RoboDK station: T1-instructions.rdk

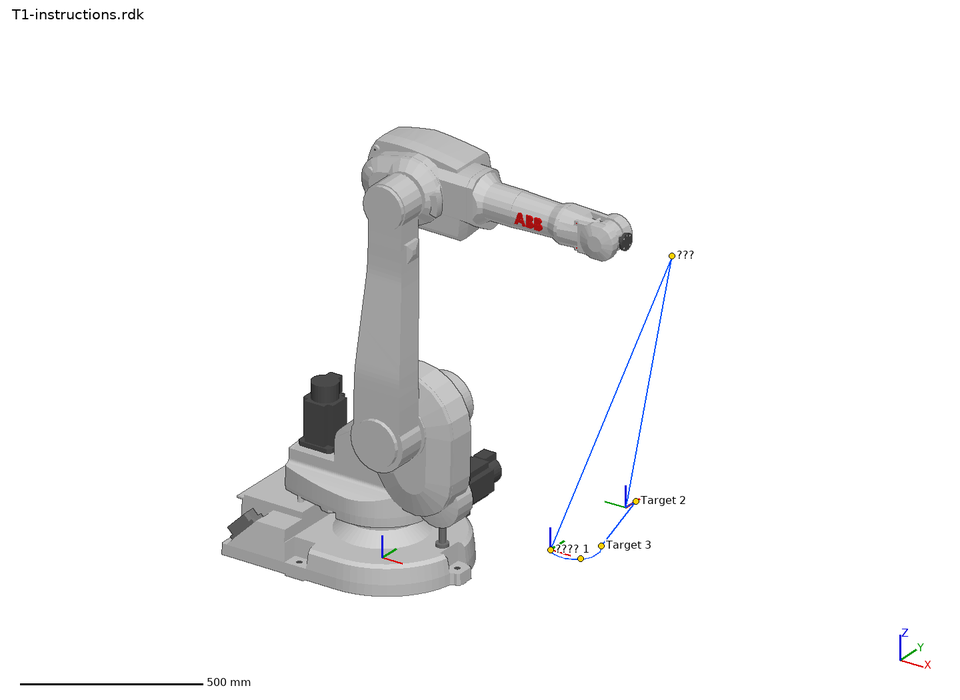
[picture v0: the station drawn from its stored meshes, robots at their saved joint values, targets as dots, program paths as lines]
Station T1 Синтетика (saved by RoboDK 5.9.4). Poses are relative to the parent item; angles as X-Y-Z fixed-axis rotations.
Station parameters (name, value as stored): T1_PARAM, 42
  - frame ABB IRB 1600-6/1.45 Base at (0, 0, 0) mm
    - robot ABB IRB 1600-6/1.45: 6 axes, payload 6 kg, reach 1450 mm, repeatability 0.05 mm, weight 250 kg
        modified DH rows (alpha deg, a mm, theta deg, d mm): 0, 0, 0, 486.5; -90, 150, -90, 0; 0, 700, 0, 0; -90, 0, 0, 600; 90, 0, 0, 0; -90, 0, 180, 65
        joint limits [-180, -90, -245, -200, -115, -400] to [180, 120, 65, 200, 115, 400]; home [0, 0, 0, 0, 0, 0]; saved at [0, 0, 0, 0, 0, 0]
      - tool , TCP at (0, 0, 150) mm, rotated rx 0 ry 30 rz 0 deg
  - frame Рамка 1 at (700, -200, 300) mm
    - target Дом (joint target) at (265, 200, 886.5) mm, rotated rx -180 ry 60 rz -180 deg; joints [0, 10, 10, 0, 40, 0] of ABB IRB 1600-6/1.45
    - target Цель 1 (Cartesian target) at (0, 0, 0) mm, rotated rx 180 ry 0 rz 0 deg; joints [0, 0, 0, 0, 0, 0] of ABB IRB 1600-6/1.45
    - target Target 2 (Cartesian target) at (100, 0, 0) mm, rotated rx 180 ry 0 rz 0 deg; joints [0, 0, 0, 0, 0, 0] of ABB IRB 1600-6/1.45
    - target Target 3 (Cartesian target) at (100, 100, 0) mm, rotated rx 180 ry 0 rz 0 deg; joints [0, 0, 0, 0, 0, 0] of ABB IRB 1600-6/1.45
  - frame Frame B at (600, 300, 200) mm, rotated rx 0 ry 0 rz 90 deg
    - target Target 2 (Cartesian target) at (50, 0, 0) mm, rotated rx 180 ry 0 rz 0 deg; joints [-41.186, -16.956, 4.401, -79.23, 50.002, 73.515] of ABB IRB 1600-6/1.45
  - Python program ПитонПрог (listed below)
  - program Подпрограмма (1 instructions, listed below)
  - program Программа (29 instructions, listed below)
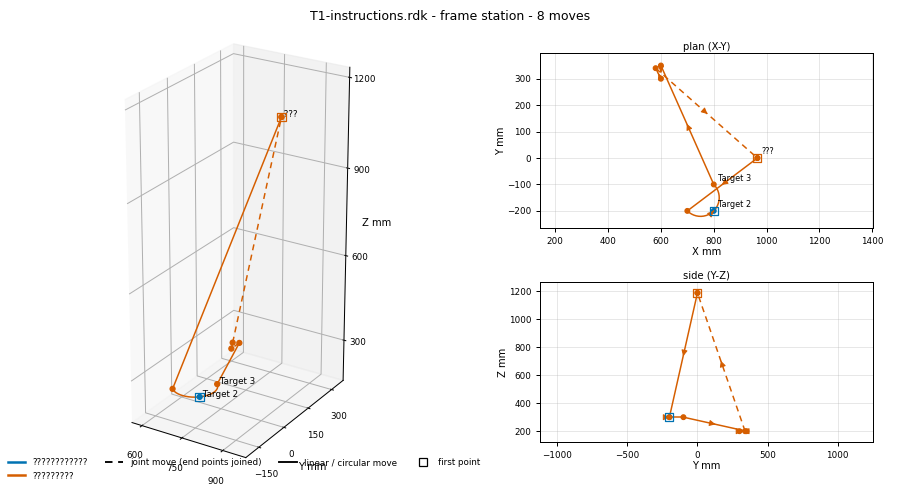
[picture p0: tool path of T1-instructions.rdk in frame station, 8 of 8 moves have a stored position in this frame; points joined in program order, loops and branches not executed]

--- Python program ПитонПрог ---
# Скрипт станции
from robodk.robolink import *
RDK = Robolink()
print("hello")

--- program Подпрограмма (robot ABB IRB 1600-6/1.45) ---
  MoveL (Target 2)

--- program Программа (robot ABB IRB 1600-6/1.45) ---
  Set Ref.: Рамка 1
  Set Tool: Инструмент 1 at (0, 0, 150) mm, rotated rx 0 ry 30 rz 0 deg
  Set speed (150.0 mm/s)
  Smooth(5)
  MoveJ (Дом)
  MoveL (Цель 1)
  MoveC (Target 2, Target 3)
  Pause 500 ms
  Stop
  Set DO_5=1
  Set AO_1=2.5
  Wait DI_3=1 T2.0s
  Wait DI_4=0
  Call SetRPM(70)
  Call Подпрограмма
  Run Подпрограмма
  Call ПитонПрог
  LaserOn
  Комментарий
  Print: Hello operator
  Set Ref.: Frame B
  MoveL (Target 2)
  MoveJ 22 to (0, 0, 0) mm; joints [10, -10, 20, 0, 40, 0]
  MoveL 23 to (40, 20, 0) mm, rotated rx 180 ry 0 rz 0 deg; joints [168.009, -54.839, -167.411, -6.113, -77.276, -9.071]
  Accurate (rounding -1 mm)
  Set speed (45.0 deg/s)
  Set accel. (200.0 deg/s2)
  Set accel. (800.0 mm/s2)
  MoveJ (Дом)
